Fanuc KAREL source: kt00033.KL

-- PROVISIONAL review KL for V1013-1; original PC SHA256 527031c7a9c61ce8ae343c1d479cea4dc6e51c0c13938546577b88ac9532c22b
-- Incomplete behavior may be omitted. Consult companion uncertainty JSON. Do not deploy.
PROGRAM KT00033
%NOLOCKGROUP
VAR
  I1 : INTEGER
  I2 : INTEGER
  OUT : INTEGER
BEGIN
  -- UNRESOLVED_PC offsets 5-16; opcodes 2E,23
  -- UNRESOLVED_PC offsets 21-32; opcodes 2E,23
  -- UNRESOLVED_PC offsets 37-48; opcodes 2E,23
  -- UNRESOLVED_PC offsets 53-64; opcodes 2E,23
  -- UNRESOLVED_PC offsets 69-88; opcodes 21,21,53,23
  -- UNRESOLVED_PC offsets 93-97; opcodes 7F
END KT00033
